TYPE ST_Tank_CIP :
STRUCT
END_STRUCT
END_TYPE

(* stored: Version 1.1.0.1, ProductVersion 3.1.4024.12
   DUT ST_Tank_CIP: Id {83c824ad-d876-40bc-80d9-ffc1eddf2012} *)
